(* IEC 61131-3 sources: avi-aoi-management/scripts/ai-eval/ngau-nhien/kho/st-ud2-den-giao-thong/khung/src, 2 files *)

(* ---- DenGiaoThong.st ---- *)
FUNCTION_BLOCK DenGiaoThong
VAR_INPUT
    NUT_NGUOI : BOOL;
    NHAP_NHAY_VANG : BOOL;
    T_XANH_MIN : TIME;
    T_VANG : TIME;
    T_NGUOI : TIME;
    T_DO_CHUNG : TIME;
    T_NHAY : TIME;
END_VAR
VAR_OUTPUT
    XE_XANH : BOOL;
    XE_VANG : BOOL;
    XE_DO : BOOL;
    NG_XANH : BOOL;
    NG_DO : BOOL;
    TRANG_THAI : INT;
END_VAR
    (* TODO: cài đặt theo đề bài *)
    XE_XANH := FALSE;
END_FUNCTION_BLOCK

(* ---- NhapNhay.st ---- *)
FUNCTION_BLOCK NhapNhay
VAR_INPUT
    EN : BOOL;
    T_NUA : TIME;
END_VAR
VAR_OUTPUT
    Q : BOOL;
END_VAR
    (* TODO: cài đặt theo đề bài *)
    Q := FALSE;
END_FUNCTION_BLOCK
